FUNCTION_BLOCK ActivePhaseAborted (* Basic Function Block Type *)
  (* Standard: 61499-2 *)
  (* Version 0.0, 10/12/2026, Schneider Electric, Template *)
  PACKAGE SE.Nereda;
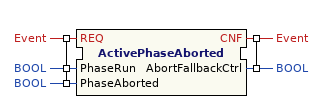
  EVENT_INPUT
    REQ WITH PhaseRun, PhaseAborted; (* Normal Execution Request *)
  END_EVENT
  EVENT_OUTPUT
    CNF WITH AbortFallbackCtrl; (* Execution Confirmation *)
  END_EVENT
  VAR_INPUT
    PhaseRun : BOOL;
    PhaseAborted : BOOL;
  END_VAR
  VAR_OUTPUT
    AbortFallbackCtrl : BOOL; (* Output event qualifier *)
  END_VAR
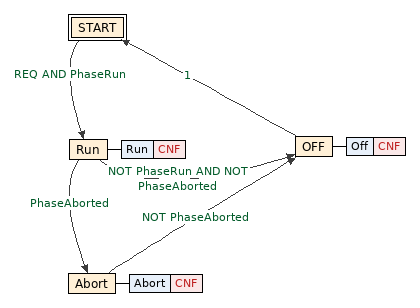
  EC_STATES
    START; (* Initial State *)
    Run : Run -> CNF; (* Normal execution *)
    Abort : Abort -> CNF;
    OFF : Off -> CNF;
  END_STATES
  EC_TRANSITIONS
    START TO Run := REQ AND PhaseRun;
    Run TO Abort := PhaseAborted;
    Run TO OFF := NOT PhaseRun AND NOT PhaseAborted;
    OFF TO START := 1;
    Abort TO OFF := NOT PhaseAborted;
  END_TRANSITIONS
  ALGORITHM Run IN ST: (* Normally executed algorithm *)
;
AbortFallbackCtrl := FALSE;
  END_ALGORITHM
  ALGORITHM Off IN ST:
;
AbortFallbackCtrl := FALSE;
  END_ALGORITHM
  ALGORITHM Abort IN ST:
;
AbortFallbackCtrl := TRUE;
  END_ALGORITHM
END_FUNCTION_BLOCK
